// // MIGRATION DRAFT: not included in PLC compilation.
// // Reference: Reference_Project/MQTT_Handler_FB.scl, object MQTT_Handler_FB.
// // Types, globals, calls, units and behavior require manual reconciliation.
// // See docs/TIA_Missing_Blocks.md before importing as PLC code.
FUNCTION_BLOCK MQTT_Handler_FB
// 
//    VAR_INPUT
//       Enable : Bool := True;
//    END_VAR
// 
//    VAR_IN_OUT
//       LMQTT_DB : LMQTT_DB_UDT;
//    END_VAR
// 
//    VAR
//       MQTT_Setup : Bool;
//       MQTT_Topic : WString;
//       Publish_Msg_Payload : Array[1..128] of Byte;
//       Received_Topic : WString;
//       Received_Msg_Payload : Array[0..1024] of Byte;
//       i : UInt;
//       j : UInt;
//       Subscribe : Bool;
//       Unsubscribe : Bool;
//       Received_Msg_Status : USInt;
//       Received_Msg_Length : UDInt;
//       Busy : Bool;
//       Valid : Bool;
//       Done : Bool;
//       Error : Bool;
//       Status : Word;
//       Diagnostics : typeDiagnostics;
//       JSON_Tree   : Array[1..18] of LStream_typeElement;
//       Shuttle_No : UInt;
//       sSubTopic : Array[1..24] of String;
//       bSubscribed : Bool;
//       SubscribeState : Int;
//       SubscribeIndex : Int := 1;
//       SubscribeCount : UInt := 1;
//       SubscribeTopicList : Array[1..30] of String;
//       sPayloadRcv : String;
//       sPayloadRcv_1 : String;
//       sPayloadRcv_2 : String;
//       sPayloadRcv_3 : String;
//       sPayloadRcv_4 : String;
//       sPayloadRcv_5 : String;
//       MQTT_AutoReset : UInt;
//       Enable_AutoReset : Bool;
//       T_AutoReset   : TON;
//    END_VAR
// 
//    VAR_TEMP
//       iIndex : UInt;
//       sIndexStr : String;
//       k : UInt;
//       test : DWord;
//       Y : UInt;
//    END_VAR

// // MIGRATION DRAFT: not included in PLC compilation.
// // Reference: Reference_Project/MQTT_Handler_FB.scl, object MQTT_Handler_FB.
// // Types, globals, calls, units and behavior require manual reconciliation.
// // See docs/TIA_Missing_Blocks.md before importing as PLC code.
// (*
// 	TODO
// 	1. Add timeout on subscribe event
// 	2. Add cyclic checks for all the different errors in the status word
// 
// 	Status word values:
// 	16#0000 Last job (publish/subscribe/unsubscribe) successfully executed
// 	16#7000 Block is idle/client not connected
// 	16#7001 First call after enable = TRUE
// 	16#7002 Block processes job
// 	16#7003 Establishing connection to MQTT broker
// 	16#7004 MQTT client connected and ready for job
// 	16#7005 Ping is sent to the broker
// 	16#7006 Publish job is executed
// 	16#7008 Subscribe job is executed
// 	16#7010 Unsubscribe job is executed
// 	*)
// 
// 	IF FirstScan THEN
// 	    MQTT_Enable := TRUE;
// 	END_IF;
// 
// 	LMQTT_DB.connParam := Settings_DB.Shuttle_MQTT.MQTT_Con_Params;
// 	LMQTT_DB.clientIdentifier := Settings_DB.Shuttle_MQTT.Client_ID;
// 	LMQTT_DB.username := Settings_DB.Shuttle_MQTT.Username;
// 	LMQTT_DB.password := Settings_DB.Shuttle_MQTT.Password;
// 	LMQTT_DB.willtopic := Settings_DB.Shuttle_MQTT.Will_Topic;
// 	LMQTT_DB.willMsgPayload := Settings_DB.Shuttle_MQTT.Will_Msg_Payload;
// 	LMQTT_DB.willMsgLen := 0;
// 	LMQTT_DB.willMsgPayload := Publish_Msg_Payload;
// 	Received_Topic := LMQTT_DB.receivedTopic;
// 	Received_Msg_Payload := LMQTT_DB.receivedMsgPayload;
// 	Received_Msg_Status:=LMQTT_DB.receivedMsgStatus;
// 	Received_Msg_Length := LMQTT_DB.receivedMsgDataLen;
// 	LMQTT_DB.enable := Enable;
// 
// 	LMQTT_DB.qos := Settings_DB.Shuttle_MQTT.QoS;
// 	LMQTT_DB.retain := Settings_DB.Shuttle_MQTT.Retain;
// 	Status := LMQTT_DB.status;
// 
// 	IF NOT bSubscribed THEN
// 	    FOR Shuttle_No := 1 TO Settings_DB.System.Shuttle_Count DO
// 	        iIndex := Shuttle_No;
// 	        sIndexStr := RemovePlusSign(UINT_TO_STRING(iIndex));
// 
// 	        sSubTopic[Shuttle_No] := CONCAT(IN1 := 'vehicle/', IN2 := 'Shuttle-');
// 	        IF iIndex < 10 THEN
// 	            sSubTopic[Shuttle_No] := CONCAT(IN1 := sSubTopic[Shuttle_No], IN2 := '0');
// 	        END_IF;
// 	        sSubTopic[Shuttle_No] := CONCAT(IN1 := sSubTopic[Shuttle_No], IN2 := sIndexStr);
// 	        sSubTopic[Shuttle_No] := CONCAT(IN1 := sSubTopic[Shuttle_No], IN2 := '/state');
// 	    END_FOR;
// 
// 	    SubscribeCount := 1;
// 	    FOR Y := 1 TO Settings_DB.System.Shuttle_Count DO
// 	        SubscribeTopicList[SubscribeCount] := sSubTopic[Y];
// 	        IF Y < Settings_DB.System.Shuttle_Count THEN
// 	            SubscribeCount := SubscribeCount + 1;
// 	        END_IF;
// 	    END_FOR;
// 
// 	    CASE SubscribeState OF
// 	        0:
// 	            IF SubscribeIndex <= SubscribeCount THEN
// 	                LMQTT_DB.mqttTopic := STRING_TO_WSTRING(SubscribeTopicList[SubscribeIndex]);
// 	                LMQTT_DB.subscribe := TRUE;
// 	                SubscribeState := 1;
// 	            ELSE
// 	                SubscribeState := 99;
// 	            END_IF;
// 
// 	        1:
// 	            IF LMQTT_DB.done THEN
// 	                LMQTT_DB.subscribe := FALSE;
// 	                SubscribeIndex := SubscribeIndex + 1;
// 	                SubscribeState := 0;
// 	            ELSIF NOT LMQTT_DB.done AND NOT LMQTT_DB.subscribe THEN
// 	                SubscribeState := 0;
// 	            ELSIF LMQTT_DB.error THEN
// 
// 	                SubscribeState := 98;
// 	                Error_Word_1.%X2 := TRUE;
// 	            END_IF;
// 
// 	        98:
// 	            LMQTT_DB.subscribe := FALSE;
// 	            bSubscribed := FALSE;
// 
// 	            IF Reset_All THEN
// 	                SubscribeCount := 0;
// 	                SubscribeIndex := 1;
// 	                SubscribeState := 0;
// 	                Error_Word_1.%X2 := FALSE;
// 	            END_IF;
// 
// 	        99:
// 	            bSubscribed := TRUE;
// 	            LMQTT_DB.subscribe := FALSE;
// 	    END_CASE;
// 	END_IF;
// 
// 	FOR k := 1 TO Settings_DB.System.Shuttle_Count DO
// 	    IF LMQTT_DB.receivedTopic = STRING_TO_WSTRING(sSubTopic[k]) THEN
// 	        sPayloadRcv := ByteArrayToString(ByteArray := LMQTT_DB.receivedMsgPayload,
// 	                                            Lenght := UDINT_TO_INT(LMQTT_DB.receivedMsgDataLen),
// 	                                            ByteArrayToString_1 => sPayloadRcv_1,
// 	                                            ByteArrayToString_2=>sPayloadRcv_2,
// 	                                            ByteArrayToString_3=>sPayloadRcv_3,
// 	                                            ByteArrayToString_4=>sPayloadRcv_4,
// 	                                            ByteArrayToString_5=>sPayloadRcv_5);
// 
// 	        IF sPayloadRcv <> '' THEN
// 	            Shuttle_MQTT_DB.Shuttle_MQTT[k].Message.Shuttle_Status := ParseShuttle_Status(String_1 := sPayloadRcv,
// 	                                                                                          String_2 := sPayloadRcv_1,
// 	                                                                                          String_3 := sPayloadRcv_2,
// 	                                                                                          String_4:=sPayloadRcv_3,
// 	                                                                                          String_5:=sPayloadRcv_4,
// 	                                                                                          String_6:=sPayloadRcv_5);
// 	        END_IF;
// 	   END_IF;
// 	END_FOR;
// 
// 	    IF Error THEN
// 
// 	        IF Status = 16#8001 THEN
// 	            Error := 0;
// 
// 	        ELSIF Status = 16#8200 THEN
// 	            Error := 0;
// 
// 	        ELSIF Status = 16#8201 THEN
// 	            Error := 0;
// 
// 
// 
// 	        ELSIF Status = 16#8210 THEN
// 	            Error := 0;
// 
// 	        ELSIF Status = 16#8220 THEN
// 	            Error := 0;
// 
// 	        ELSIF Status = 16#8230 THEN
// 	            Error := 0;
// 
// 	        ELSIF Status = 16#8300 THEN
// 	            Error := 0;
// 
// 	        ELSIF Status = 16#8310 THEN
// 	            Error := 0;
// 
// 	        ELSIF Status = 16#8320 THEN
// 	            Error := 0;
// 
// 	        ELSIF Status = 16#8600 THEN
// 	            Error := 0;
// 
// 
// 
// 	        ELSIF Status = 16#8601 THEN
// 	            Error := 0;
// 
// 	        ELSIF Status = 16#8620 THEN
// 	            Error := 0;
// 
// 	        ELSIF Status = 16#8650 THEN
// 	            Error := 0;
// 
// 	        ELSIF Status = 16#8670 THEN
// 	            Error := 0;
// 
// 	        ELSIF Status = 16#8700 THEN
// 	            Error := 0;
// 
// 	        ELSIF Status = 16#8710 THEN
// 	            Error := 0;
// 
// 	        ELSIF Status = 16#8720 THEN
// 	            Error := 0;
// 	        ELSE
// 	            ;
// 	        END_IF;
// 	    END_IF;
// 
// 	IF Reset_All THEN
// 	    SubscribeCount := 0;
// 	    SubscribeIndex := 1;
// 	    SubscribeState := 0;
// 	    bSubscribed := FALSE;
// 	END_IF;
// 
// 
// 	IF LMQTT_DB.enable AND NOT LMQTT_DB.valid AND NOT LMQTT_DB.done AND NOT LMQTT_DB.busy AND LMQTT_DB.error THEN
// 	    Enable_AutoReset := TRUE;
// 	ELSE
// 	    Enable_AutoReset := FALSE;
// 	    MQTT_AutoReset := 0;
// 	    R_Reset_All_False(CLK:=TRUE);
// 	    IF R_Reset_All_False.Q THEN
// 	        Reset_All := FALSE;
// 	    END_IF;
// 	END_IF;
// 
// 	IF Enable_AutoReset THEN
// 	    CASE MQTT_AutoReset OF
// 	        0:
// 	            MQTT_AutoReset := MQTT_AutoReset + 1;
// 	        1:
// 	            LMQTT_DB.enable := FALSE;
// 	            MQTT_AutoReset := MQTT_AutoReset + 1;
// 	        2:
// 	            Reset_All := TRUE;
// 	            MQTT_AutoReset := MQTT_AutoReset + 1;
// 	        3:
// 	            T_AutoReset(IN:=TRUE,
// 	                         PT:=t#10s);
// 	            IF T_AutoReset.Q THEN
// 	                T_AutoReset(IN := FALSE,
// 	                             PT := t#0s);
// 	                             Reset_All := FALSE;
// 	                MQTT_AutoReset := MQTT_AutoReset + 1;
// 	            END_IF;
// 
// 	        4:
// 	            LMQTT_DB.enable := TRUE;
// 	            MQTT_AutoReset := MQTT_AutoReset + 1;
// 
// 	        5:
// 	            IF LMQTT_DB.enable AND NOT LMQTT_DB.valid AND NOT LMQTT_DB.done AND NOT LMQTT_DB.busy AND LMQTT_DB.error THEN
// 	                T_AutoReset(IN := TRUE,
// 	                             PT := t#3s);
// 
// 	                IF T_AutoReset.Q THEN
// 	                    MQTT_AutoReset := 1;
// 	                END_IF;
// 	            END_IF;
// 
// 
// 	    END_CASE;
// 	END_IF;

END_FUNCTION_BLOCK

(* stored: Version 1.1.0.1
   POU MQTT_Handler_FB: Id {f6b145c9-8e64-5184-94aa-af1ffe4243d4}, SpecialFunc None *)
